(* IEC 61131-3 sources: nautilus/siemens/writer/testdata/pous, 2 files *)

(* ---- lib.st ---- *)
(* The library of the project's-blocks fixture (#1301): global constants,
   two FUNCTIONs and two FUNCTION_BLOCKs, one inside the other. *)
VAR_GLOBAL CONSTANT
    HI_LIMIT : REAL := 80.0;
    T_DELAY  : TIME := T#30ms;
    STEPS    : INT := 3;
    LOW      : INT := -2;
END_VAR

FUNCTION Scale : REAL
VAR_INPUT
    Raw : REAL;
    Lo  : REAL;
    Hi  : REAL;
END_VAR
VAR
    span : REAL;
END_VAR
span := Hi - Lo;
IF span <= 0.0 THEN
    Scale := Lo;
    RETURN;
END_IF;
Scale := Lo + Raw * span / 100.0;
END_FUNCTION

FUNCTION Bump : INT
VAR_INPUT
    X : INT;
END_VAR
Bump := X + 1;
END_FUNCTION

FUNCTION_BLOCK Debounce
VAR_INPUT
    IN : BOOL;
    PT : TIME;
END_VAR
VAR_OUTPUT
    Q : BOOL;
END_VAR
VAR
    t : TON;
END_VAR
t(IN := IN, PT := PT);
Q := t.Q;
END_FUNCTION_BLOCK

FUNCTION_BLOCK Station
VAR_INPUT
    Run   : BOOL;
    Level : REAL;
END_VAR
VAR_OUTPUT
    High  : BOOL;
    Count : DINT;
    Total : INT;
END_VAR
VAR_IN_OUT
    Starts : INT;
END_VAR
VAR
    db   : Debounce;
    edge : R_TRIG;
    i    : INT;
    hold : TON;
END_VAR
VAR_TEMP
    scratch : INT := 10;
END_VAR
VAR CONSTANT
    GAIN : REAL := 2.0;
    TOP  : INT := 6;
END_VAR
db(IN := Run, PT := T_DELAY);
edge(CLK := db.Q);
IF edge.Q THEN
    Starts := Starts + 1;
    Count := Count + 1;
END_IF;
High := Level * GAIN > HI_LIMIT;
Total := 0;
FOR i := 1 TO STEPS DO
    Total := Total + i;
END_FOR;
CASE Total OF
    TOP: Total := LOW;
END_CASE;
scratch := scratch + Total;
hold(IN := High);
END_FUNCTION_BLOCK

(* ---- Main.st ---- *)
PROGRAM Main
(* Two instances of the library's Station, one bound to tags and one to a
   local; the library's FUNCTIONs in expressions, positional and formal. *)
VAR_EXTERNAL
    Run    : BOOL;
    Level  : REAL;
    Starts : INT;
    High   : BOOL;
    Pct    : REAL;
    Count  : DINT;
    Next   : INT;
END_VAR
VAR
    st1         : Station;
    st2         : Station;
    localStarts : INT;
END_VAR
st1(Run := Run, Level := Level, Starts := Starts, High => High, Count => Count);
st2(Run := NOT Run, Level := Scale(Level, 0.0, HI_LIMIT), Starts := localStarts);
Pct := Scale(Raw := Level, Lo := 0.0, Hi := 100.0);
Next := Bump(Starts) + st1.Total;
END_PROGRAM
